// GRAFCET G3 Werkstückrotation [Langfeld].
{attribute 'qualified_only'}
{attribute 'strict'}
{attribute 'to_string'}
TYPE E_G3Step :
(
    S30_Bereit := 30,
    S31_Stop := 31,     // Master steht an der Rotationsposition
    S32_Drehen := 32    // W dreht
) INT;
END_TYPE

(* stored: Version 1.1.0.1
   DUT E_G3Step: Id {0eb9916f-b4fb-52cb-8082-8ee8b8e3f604} *)
